(* IEC 61131-3 sources: volt/packages/volt-lsp-iec/test-corpus/bakon-nano/Device/Plc Logic/Application/Library Manager/L_EtcSlaveConfig, 51 files *)

(* ---- _L_ECC_ESCHEDULE.dut ---- *)
TYPE _L_ECC_ESCHEDULE :
(
	INIT := 0,
	INIT_DONE := 99,
	SCHEDULING_ACTIVE := 10
);
END_TYPE

(* ---- _L_ECC_ESEVERITY.dut ---- *)
TYPE _L_ECC_ESEVERITY :
(
	NO_RESPONSE := 0,
	WARNING := 2,
	INFORMATION := 11,
	WARNING_LOCK := 13,
	FAULT_LOG := 18,
	FAULT_QSPAPPL := 19,
	FAULT_QSP := 20,
	FAULT_QSP_CINH := 21,
	FAULT_CINH := 23,
	FAULT := 30
);
END_TYPE

(* ---- _L_ECC_ESTEPPER.dut ---- *)
TYPE _L_ECC_ESTEPPER :
(
	INIT := 0,
	INIT_DONE := 99,
	READ_IDENTITY_INIT := 10,
	READ_IDENTITY_DEVICENAME,
	READ_IDENTITY_HARDWAREVERSION,
	READ_IDENTITY_SOFTWAREVERSION,
	READ_IDENTITY_SYSTEMVERSION,
	READ_IDENTITY_VENDORID,
	READ_IDENTITY_PRODUCTCODE,
	READ_IDENTITY_REVISION,
	READ_IDENTITY_SERIALNUMBER,
	READ_IDENTITY_MANUFACTURER,
	READ_IDENTITY_DEVICECLASS,
	READ_IDENTITY_PRODUCTCODE_CD,
	READ_IDENTITY_FINISH_CD,
	C250_INIT := 100,
	C250_ERROR_REGISTER := 110,
	C250_CHECK_READING_REQUIRED,
	C250_EXTERNAL_TEMPERATURE := 115,
	C250_STATE_INPUTS,
	C250_STATE_OUTPUTS,
	C250_CPU1_REFERENCE_VOLTAGE := 120,
	C250_CPU1_24V_VOLTAGE := 121,
	C250_CPU1_5V_VOLTAGE := 122,
	C250_CPU1_3V3_VOLTAGE := 123,
	C250_CPU1_TEMPERATURE := 124,
	C250_CPU1_OUTPUT_CURRENT := 125,
	C250_CPU1_CYCLETIME := 126,
	C250_CPU1_ERROR_CODE := 127,
	C250_CPU1_ERROR_LINE := 128,
	C250_CPU1_ERROR_MODULE := 129,
	C250_CPU1_ERROR_CLASS := 130,
	C250_CPU1_ERROR_WRITETOCONTROLLER := 131,
	C250_CPU1_ERROR_WRITETOFRAMEWORK := 132,
	C250_CPU2_REFERENCE_VOLTAGE := 140,
	C250_CPU2_24V_VOLTAGE,
	C250_CPU2_5V_VOLTAGE,
	C250_CPU2_3V3_VOLTAGE,
	C250_CPU2_TEMPERATURE,
	C250_CPU2_OUTPUT_CURRENT,
	C250_CPU2_CYCLETIME,
	C250_CPU2_ERROR_CODE,
	C250_CPU2_ERROR_LINE,
	C250_CPU2_ERROR_MODULE,
	C250_CPU2_ERROR_CLASS,
	C250_CPU2_ERROR_WRITETOCONTROLLER,
	C250_CPU2_ERROR_WRITETOFRAMEWORK := 152,
	C250_DONE_WRITETOLOGS := 198,
	C250_DONE := 199,
	S13X_INIT := 200,
	S13X_DISABLE_AUTO_ACK,
	S13X_ERROR_REGISTER_HARDWARE := 210,
	S13X_ERROR_REGISTER_DIAGNOSTIC,
	S13X_MODULE_STATUS_DIAGNOSTIC,
	S13X_CHECK_READING_REQUIRED,
	S13X_COUPLER_VERSION_FPGA := 220,
	S13X_COUPLER_VERSION_BACKPLANE,
	S13X_COUPLER_VERSION_FIRMWARE,
	S13X_COUPLER_MX_FILE,
	S13X_COUPLER_NUMBER_OF_SLICES,
	S13X_SLICE_INIT := 230,
	S13X_SLICE_VERSION_FPGA,
	S13X_SLICE_VERSION_MODULE,
	S13X_SLICE_SERIALNUMBER,
	S13X_SLICE_MX_FILE,
	S13X_SLICE_ID_CONFIGURED,
	S13X_SLICE_ADDRESS,
	S13X_SLICE_ID_DETECTED,
	S13X_SLICE_DONE,
	S13X_SLICE_SW_VERSION,
	S13X_SLICE_HW_VERSION,
	S13X_SLICE_MODULE_ID,
	S13X_SLICE_ERROR_HARDWARE_SLOT := 250,
	S13X_SLICE_ERROR_HARDWARE_DIAG1,
	S13X_SLICE_ERROR_HARDWARE_DIAG2,
	S13X_SLICE_ERROR_HARDWARE_DIAG3,
	S13X_SLICE_ERROR_HARDWARE_DIAG4,
	S13X_SLICE_ERROR_HARDWARE_WRITE_ACK,
	S13X_SLICE_ERROR_HARDWARE_WRITETOCONTROLLER,
	S13X_SLICE_ERROR_HARDWARE_WRITETOFRAMEWORK,
	S13X_SLICE_ERROR_DIAGNOSTIC_READSLOT,
	S13X_SLICE_ERROR_DIAGNOSTIC_WRITESLOT,
	S13X_SLICE_ERROR_DIAGNOSTIC_DIAG1,
	S13X_SLICE_ERROR_DIAGNOSTIC_DIAG2,
	S13X_SLICE_ERROR_DIAGNOSTIC_DIAG3,
	S13X_SLICE_ERROR_DIAGNOSTIC_DIAG4,
	S13X_SLICE_ERROR_DIAGNOSTIC_WRITE_ACK,
	S13X_SLICE_ERROR_DIAGNOSTIC_WRITETOCONTROLLER,
	S13X_SLICE_ERROR_DIAGNOSTIC_WRITETOFRAMEWORK,
	S13X_DONE_WRITETOLOGS := 298,
	S13X_DONE := 299,
	ISERIES_INIT := 400,
	ISERIES_STEP_1 := 401,
	ISERIES_STEP_2 := 402,
	ISERIES_STEP_3 := 403,
	ISERIES_STEP_4 := 404,
	ISERIES_STEP_5 := 405,
	ISERIES_DONE := 499
);
END_TYPE

(* ---- FILE_STATE.dut ---- *)
TYPE FILE_STATE :
(
	S_NONE,
	S_INITIALIZE,
	S_GET_SLAVE_STATE,
	S_WAIT_FILE_SIZE,
	S_WAIT_FILE_OPEN,
	S_READ_FILE,
	S_CLOSE_FILE,
	S_PROCESS,
	S_READ_PAR_RECORDS,
	S_WAIT_XFER_COMPLETE,
	S_ERROR,
	S_DONE
);
END_TYPE

(* ---- L_ECC_EC250_CPUNUMBER.dut ---- *)
TYPE L_ECC_EC250_CPUNUMBER :
(
	NO_CPU := 0,
	CPU_1 := 1,
	CPU_2 := 2,
	CPU_3 := 3
);
END_TYPE

(* ---- L_ECC_EC250_ERRORCLASS.dut ---- *)
TYPE L_ECC_EC250_ERRORCLASS :
(
	NO_ERROR := 0,
	SYNCHRONIZATION_ERROR := 1,
	COMMUNICATION_ERROR := 2,
	IO_ERROR := 3,
	ERRORHANDLER_ERROR := 4,
	FATAL_ERROR := 5
);
END_TYPE

(* ---- L_ECC_EC250_ERRORCODE.dut ---- *)
TYPE L_ECC_EC250_ERRORCODE :
(
	OK := 0,
	HWT_PARAMETER_ERROR := 1,
	HWT_INIT_ERROR := 2,
	HWT_MEM_MARCHC_ERROR := 100,
	HWT_MEM_GALPAT_ERROR := 101,
	HWT_STACK_UNDERFLOW_ERROR := 200,
	HWT_STACK_OVERFLOW_ERROR := 201,
	HWT_CPU_ERROR := 300,
	WT_FW_ERROR := 400,
	HWT_FWINTERFACE_ERROR := 500,
	HWT_ADC_ERROR := 504,
	HWT_DMA_ERROR := 505,
	HWT_CRC_ERROR := 506,
	HWT_TIMER_ERROR := 507,
	HWT_CLOCK_ERROR := 508,
	HWT_SOFTERROR := 509,
	HWT_DIVZERO := 510,
	TIMEOUT_ERR := 512,
	OUT_OF_RANGE_ERR := 513,
	OVERWRITE_ERR := 514,
	UNDERFLOW_ERR := 515,
	PRG_CNTRL_ERR := 516,
	INIT_ERROR := 528,
	ASSERT_TRUE_ERR := 592,
	ASSERT_NOT_NULL_ERR := 593,
	ASSERT_GE_ERR := 594,
	ASSERT_GT_ERR := 595,
	ASSERT_LE_ERR := 596,
	ASSERT_LT_ERR := 597,
	ASSERT_NE_ERR := 598,
	ASSERT_EQ_ERR := 599,
	ASSERT_FALSE_ERR := 600,
	TP_OUT_NOT_SPECIFIED := 640,
	TP_OUT_NOT_RECOGNIZED := 641,
	TP_OUT_NOT_ACTIVE := 642,
	TP_INP_BUSY := 656,
	TP_INP_CROSSTALK := 657,
	TP_INP_NOT_RECOGNIZED := 658,
	TP_INTINP_NOT_RECOGNIZED := 659,
	TP_INP_LOST := 660,
	TP_INVALID_COUNT_FOR_SELECTOR := 661,
	MRAM_READ_ERR := 673,
	MRAM_WRITE_ERR := 674,
	MRAM_INDEX_OUT_OF_RANGE := 675,
	MRAM_CORRUPT_PAGE_SIZE := 676,
	MRAM_CRC_ERR := 677,
	MRAM_MAGICNUMBER_ERR := 678,
	RESET_LOW_POWER := 768,
	RESET_WINDOW_WD := 769,
	RESET_INDEPENDENT_WD := 770,
	RESET_SW := 771,
	RESET_POWER_ON_DOWN := 772,
	RESET_NMI := 773,
	RESET_BROWNOUT := 774,
	RESET_NO_REASON := 775,
	ADC_REF_LOW := 1024,
	ADC_REF_HIGH := 1025,
	ADC_24V_LOW := 1026,
	ADC_24V_HIGH := 1027,
	ADC_5V_LOW := 1028,
	ADC_5V_HIGH := 1029,
	ADC_3_3V_LOW := 1030,
	ADC_3_3V_HIGH := 1031,
	ADC_TEMP_LOW := 1032,
	ADC_TEMP_HIGH := 1033,
	ADC_CURR_HIGH := 1034,
	ADC_24V_FATAL := 1035,
	LINE_TIMEOUT := 1280,
	NOVALIDCPUID := 1281,
	TIMEOUTTIMERERR := 1282,
	DIPSWITCHREADERR := 1283,
	DIPSWITCHCHANGED := 1284,
	DIPSWITCHXCHGERROR := 1285,
	DIPSWITCH_INVALID_ADDRESS := 1286,
	CLK_ERROR := 1312,
	CLK_PARTNER_LOW := 1313,
	CLK_PARTNER_HIGH := 1314,
	HW_REVISION_ERROR := 1328,
	INPUTXCHGERROR := 1536,
	INPUT_TIMEOUT := 1537,
	INPUT_EXTMATTE_KS := 1552,
	INPUT_EXTMATTE_OPEN := 1553,
	OUTPUTXCHGERROR := 1792,
	OUTPUTFAIL := 1793,
	OUTPUT_WAITFB := 1794,
	OUTPUT_TIMEOUT := 1795,
	OUTPUT_HSTP_TIMEOUT := 1796,
	OUTPUT_LSTP_TIMEOUT := 1797,
	OUTPUT_LSTP_CONNECT_ERR := 1798,
	OUTPUT_USTP_TIMEOUT := 1799,
	OUTPUT_NOPAR_USED := 1800,
	BCOM_NOTREADY := 2048,
	BCOM_BUSY := 2049,
	BCOM_NONEWDATA := 2050,
	BCOM_CRCERR := 2051,
	BCOM_BITERR := 2052,
	XCOM_NOTREADY := 2304,
	XCOM_BUSY := 2305,
	XCOM_NONEWDATA := 2306,
	XCOM_CRCERR := 2307,
	I2C_TIMEOUT := 2560,
	I2C_BUSY := 2561,
	FSOE_RESET_IND := 2816,
	FSOE_INVALID_CMD := 2817,
	FSOE_UNKNOWN_CMD := 2818,
	FSOE_INVALID_CONNID := 2819,
	FSOE_INVALID_CRC := 2820,
	FSOE_WD_EXPIRED := 2821,
	FSOE_INVALID_ADDRESS := 2822,
	FSOE_INVALID_DATA := 2823,
	FSOE_INVALID_COMMPARALEN := 2824,
	FSOE_INVALID_COMMPARA := 2825,
	FSOE_INVALID_USERPARALEN := 2826,
	FSOE_INVALID_USERPARA := 2827,
	FSOE_INVALID_TP_INP_DURATION := 2828,
	FSOE_INVALID_TP_INP_FREQUENCY := 2829,
	FSOE_INVALID_TP_OUT_DURATION := 2830,
	FSOE_INVALID_TP_OUT_FREQUENCY := 2831,
	FSOE_INVALID_WATCHDOG_TIME := 2832,
	FSOE_INVALID_INP_EXT_SUPPLY := 2833,
	FSOE_INVALID_INP_IN_USE := 2834,
	FSOE_INVALID_INP_USED_EXT_MISMATCH := 2835,
	FSOE_INVALID_OUT_IN_USE := 2836,
	FSOE_INVALID_OUT_USED_EXT_MISMATCH := 2837,
	FSOE_EXTENDED_ERROR := 2944,
	FSOE_ERROR := 2992,
	TH_GLOBAL_ERROR := 3072,
	TH_TIMEOUT := 3073,
	MC1_ID_INVALID := 3329,
	MC2_ID_INVALID := 3330,
	MC3_ID_INVALID := 3331,
	FOREIGN_ERROR_DETECTED := 3584,
	FLASH_TIMEOUT := 3841,
	FLASH_LOCKED := 3842,
	FLASH_BUSY := 3851,
	FLASH_ERROR := 3854
);
END_TYPE

(* ---- L_ECC_EC250_ERRORMODULE.dut ---- *)
TYPE L_ECC_EC250_ERRORMODULE :
(
	OBJ_UNKNOWN_ID := 0,
	OBJ_FSOETASK_ID := 4,
	OBJ_INPUT_ID := 8,
	OBJ_MAINTASK_ID := 12,
	OBJ_PRGCONTRLTASK_ID := 16,
	OBJ_SYNCSAFETYPARTNER_ID := 20,
	OBJ_XCOM_ID := 24,
	OBJ_SAFETYHAL_ID := 28,
	OBJ_YSTIMER_ID := 32,
	OBJ_MSTIMER_ID := 36,
	OBJ_BASEBOARDCOM_ID := 44,
	OBJ_DIPSWITCH_ID := 48,
	OBJ_HELPER_ID := 52,
	OBJ_SYNCLINE_ID := 56,
	OBJ_TIMETABLE_ID := 60,
	OBJ_TESTHANDLER_ID := 64,
	OBJ_TIME_ITERATOR_ID := 80,
	OBJ_SPI_ID := 96,
	OBJ_TIMER_ID := 97,
	OBJ_BACKUPSRAM_ID := 98,
	OBJ_PWR_ID := 99,
	OBJ_RCC_ID := 100,
	OBJ_GPIO_ID := 101,
	OBJ_DMASTREAM_ID := 102,
	OBJ_ADC_ID := 103,
	OBJ_WD_ID := 104,
	OBJ_FLASH_ID := 105,
	OBJ_I2C_ID := 106,
	OBJ_INPUTHANDLER_ID_1 := 128,
	OBJ_INPUTHANDLER_ID_2 := 129,
	OBJ_INPUTHANDLER_ID_3 := 130,
	OBJ_INPUTHANDLER_ID_4 := 131,
	OBJ_OUTPUT_ID_1 := 144,
	OBJ_OUTPUT_ID_2 := 145,
	OBJ_USTESTPULSE_ID := 148,
	OBJ_OUTPUTHANDLER_ID := 160,
	OBJ_OUTPFSWITCH_ID := 164
);
END_TYPE

(* ---- L_ECC_EDEVICETYPE.dut ---- *)
TYPE L_ECC_EDEVICETYPE :
(
	UNKNOWN := 0,
	C25BAYCB := 16#43004342,
	C25BAYSQ := 16#43005153,
	C25BAYA42 := 16#43000402,
	C25BAYA82 := 16#43000802,
	C25BAYA160 := 16#43001000,
	C25BAYA164 := 16#43001004,
	EPM_S130 := 16#514,
	EPM_S131 := 16#51E,
	EPM_S200 := 16#19F82,
	EPM_S201 := 16#39F84,
	EPM_S202 := 16#59FC1,
	EPM_S203 := 16#89F84,
	EPM_S204 := 16#29F82,
	EPM_S205 := 16#49F84,
	EPM_S206 := 16#79FC1,
	EPM_S207 := 16#F0147C1,
	EPM_S208 := 16#F0347C2,
	EPM_S209 := 16#139FC1,
	EPM_S210 := 16#121F41,
	EPM_S300 := 16#101AF90,
	EPM_S301 := 16#104AFA0,
	EPM_S302 := 16#106AFC8,
	EPM_S303 := 16#103AF90,
	EPM_S304 := 16#105AFA0,
	EPM_S305 := 16#107AFC8,
	EPM_S306 := 16#102AF90,
	EPM_S308 := 16#109AF90,
	EPM_S309 := 16#108AFA0,
	EPM_S310 := 16#F4157E1,
	EPM_S311 := 16#F4357E2,
	EPM_S312 := 16#1132F48,
	EPM_S400 := 16#40115C3,
	EPM_S401 := 16#40415C4,
	EPM_S402 := 16#40215C3,
	EPM_S403 := 16#40515C4,
	EPM_S404 := 16#4061544,
	EPM_S405 := 16#4031543,
	EPM_S406 := 16#40C1543,
	EPM_S408 := 16#40B1543,
	EPM_S409 := 16#4111543,
	EPM_S410 := 16#40715C3,
	EPM_S411 := 16#8411809,
	EPM_S412 := 16#40D1544,
	EPM_S413 := 16#4121544,
	EPM_S414 := 16#40E1544,
	EPM_S415 := 16#40F1543,
	EPM_S416 := 16#8842880,
	EPM_S500 := 16#50125D8,
	EPM_S501 := 16#50325E0,
	EPM_S502 := 16#50225D8,
	EPM_S503 := 16#50425E0,
	EPM_S504 := 16#50B25D8,
	EPM_S505 := 16#50A25E0,
	EPM_S600 := 16#8C13800,
	EPM_S601 := 16#8C3380A,
	EPM_S602 := 16#8C23801,
	EPM_S603 := 16#8C4388B,
	EPM_S604 := 16#9C17800,
	EPM_S606 := 16#8812880,
	EPM_S620 := 16#9014880,
	EPM_S640 := 16#E010700,
	EPM_S650 := 16#E411700
);
END_TYPE

(* ---- L_ECC_EEPMSXXX_ERRORCODE.dut ---- *)
TYPE L_ECC_EEPMSXXX_ERRORCODE :
(
	OK := 0,
	INTERNAL_ERROR := 1,
	EXTERNAL_ERROR := 2,
	CHANNEL_ERROR := 3,
	SUPPLY_VOLTAGE_ERROR := 4,
	PARAMETER_ERROR := 5,
	INTERNAL_COM_FAULT := 6,
	PROCESS_ALARM_LOST := 7,
	BROKEN_WIRE := 8,
	MEASURING_RANGE_UNDERFLOW := 9,
	MEASURING_RANGE_OVERFLOW := 10,
	LOST_OVERFLOW_UNDERFLOW_ALARM := 11,
	LOST_COMPARE_VALUE_RACHED_ALARM := 12,
	AUTO_ACK_DISABLED := 100
);
END_TYPE

(* ---- L_ECC_EERROR.dut ---- *)
TYPE L_ECC_EERROR :
(
	NOERROR := 0,
	NOSLAVECONNECTED,
	INVALIDSLAVECONNECTED,
	SLAVENOTREADYFORSDO,
	INVALIDSTATEMACHINE,
	INVALIDSLICENUMBER,
	COULDNOTSENDAUTOACKERROR,
	COULDNOTSENDDIAGNOSTICERROR
);
END_TYPE

(* ---- L_ECC_EEXTENDEDSTATE.dut ---- *)
TYPE L_ECC_EEXTENDEDSTATE :
(
	NONE := 16#0,
	INITIALIZING := 16#1,
	PREOPERATIONAL := 16#2,
	BOOTSTRAP := 16#3,
	SAFEOPERATIONAL := 16#4,
	OPERATIONAL := 16#8,
	UNKNOWN := 16#FFEF,
	FIRMWAREDOWNLOAD := 16#201,
	CABLENOTCONNECTED := 16#202,
	BUSMISMATCH := 16#203,
	CONNECTIONFAULTY := 16#801,
	NOTALLSLAVESOPERATIONAL := 16#802,
	CONNECTIONLOST := 16#803
);
END_TYPE

(* ---- L_ECC_SCC250_CPU.dut ---- *)
TYPE L_ECC_SCC250_CPU :
STRUCT
	ECPUNUMBER : L_ECC_eC250_CpuNumber;
	XERRORACTIVE : BOOL;
	EERRORCLASS : L_ECC_eC250_ErrorClass;
	EERRORCODE : L_ECC_eC250_ErrorCode;
	EPREVIOUSERRORCODE : L_ECC_eC250_ErrorCode;
	EERRORMODULE : L_ECC_eC250_ErrorModule;
	WERRORLINE : WORD;
END_STRUCT
END_TYPE

(* ---- L_ECC_SCDEVICEINFO.dut ---- *)
TYPE L_ECC_SCDEVICEINFO :
STRUCT
	UIDEVICEADDRESS : UINT;
	EDEVICETYPE : L_ECC_eDeviceType := L_ECC_eDeviceType.Unknown;
	SDEVICENAME : STRING(255);
	SHARDWAREVERSION : STRING(64);
	SSOFTWAREVERSION : STRING(64);
	USISYSTEMVERSION : USINT;
	DWVENDORID : DWORD;
	DWPRODUCTCODE : DWORD;
	DWREVISION : DWORD;
	DWSERIALNUMBER : DWORD;
END_STRUCT
END_TYPE

(* ---- L_ECC_SCEMPSXXX_DIAGNOSTIC.dut ---- *)
TYPE L_ECC_SCEMPSXXX_DIAGNOSTIC :
UNION
	SCEPMS404_S405 : L_ECC_scEPMS404_S405_Diagnostic;
	SCEPMS600 : L_ECC_scEPMS600_Diagnostic;
	SCEPMS601_S602 : L_ECC_scEPMS603_S604_Diagnostic;
	SCEPMS603_S604 : L_ECC_scEPMS603_S604_Diagnostic;
	SCGENERIC : L_ECC_scEMPSxxx_DiagnosticBits;
	ABYBYTES : ARRAY [1..4] OF BYTE;
	DWVALUE : DWORD;
END_UNION
END_TYPE

(* ---- L_ECC_SCEMPSXXX_DIAGNOSTICBITS.dut ---- *)
TYPE L_ECC_SCEMPSXXX_DIAGNOSTICBITS :
STRUCT
	BERROR : BIT;
	BINTERNALERROR : BIT;
	BEXTERNALERROR : BIT;
	BCHANNELERROR : BIT;
	BSUPPLYVOLTAGEERROR : BIT;
	BRESERVED_0 : BIT;
	BRESERVED_1 : BIT;
	BPARAMETERERROR : BIT;
	BRESERVED_2 : BIT;
	BRESERVED_3 : BIT;
	BRESERVED_4 : BIT;
	BRESERVED_5 : BIT;
	BINTERNALCOMFAULT : BIT;
	BRESERVED_6 : BIT;
	BPROCESSALARMLOST : BIT;
	BRESERVED_7 : BIT;
END_STRUCT
END_TYPE

(* ---- L_ECC_SCEPMS404_S405_DIAGNOSTIC.dut ---- *)
TYPE L_ECC_SCEPMS404_S405_DIAGNOSTIC :
STRUCT
	SCGENERAL : L_ECC_scEMPSxxx_DiagnosticBits;
	SCCHANNEL_0 : L_ECC_scEPMS404_S405_DiagnosticBits;
	SCCHANNEL_1 : L_ECC_scEPMS404_S405_DiagnosticBits;
END_STRUCT
END_TYPE

(* ---- L_ECC_SCEPMS404_S405_DIAGNOSTICBITS.dut ---- *)
TYPE L_ECC_SCEPMS404_S405_DIAGNOSTICBITS :
STRUCT
	BPARAMETERERROR : BIT;
	BRESERVED_0 : BIT;
	BRESERVED_1 : BIT;
	BRESERVED_2 : BIT;
	BBROKENWIRE : BIT;
	BPROCESSALARMLOST : BIT;
	BMEASURINGRANGEUNDERFLOW : BIT;
	BMEASURINGRANGEOVERFLOW : BIT;
END_STRUCT
END_TYPE

(* ---- L_ECC_SCEPMS600_DIAGNOSTIC.dut ---- *)
TYPE L_ECC_SCEPMS600_DIAGNOSTIC :
STRUCT
	SCGENERAL : L_ECC_scEMPSxxx_DiagnosticBits;
	SCCHANNEL_0 : L_ECC_scEPMS600_DiagnosticBits;
	BYRESERVED_1 : BYTE;
END_STRUCT
END_TYPE

(* ---- L_ECC_SCEPMS600_DIAGNOSTICBITS.dut ---- *)
TYPE L_ECC_SCEPMS600_DIAGNOSTICBITS :
STRUCT
	BHW_GATEOPENED : BIT;
	BHW_GATECLOSED : BIT;
	BENDVALUEOVERFLOWUNDERFLOW : BIT;
	BCOMPAREVALUEREACHED : BIT;
	BLATCHED : BIT;
	BRESERVED_0 : BIT;
	BRESERVED_1 : BIT;
	BRESERVED_2 : BIT;
END_STRUCT
END_TYPE

(* ---- L_ECC_SCEPMS601_S602_DIAGNOSTICBITS.dut ---- *)
TYPE L_ECC_SCEPMS601_S602_DIAGNOSTICBITS :
STRUCT
	BRESERVED_0 : BIT;
	BLOSTOVERFLOWUNDERFLOWALARM : BIT;
	BLOSTCOMPAREVALUEREACHEDALARM : BIT;
	BRESERVED_1 : BIT;
	BRESERVED_2 : BIT;
	BRESERVED_3 : BIT;
	BRESERVED_4 : BIT;
END_STRUCT
END_TYPE

(* ---- L_ECC_SCEPMS603_S604_DIAGNOSTIC.dut ---- *)
TYPE L_ECC_SCEPMS603_S604_DIAGNOSTIC :
STRUCT
	SCGENERAL : L_ECC_scEMPSxxx_DiagnosticBits;
	BYRESERVED_0 : BYTE;
	BYRESERVED_1 : BYTE;
END_STRUCT
END_TYPE

(* ---- L_ECC_SCS13X_COUPLER.dut ---- *)
TYPE L_ECC_SCS13X_COUPLER :
STRUCT
	WNUMBEROFIOSLICES : WORD;
	UIVERSION_FPGA : UINT;
	UIVERSION_BACKPLANE : UINT;
	UDIVERSION_FIRMWARE : UDINT;
	SMX_FILE : STRING(16);
END_STRUCT
END_TYPE

(* ---- L_ECC_SCS13X_IO_SLICE.dut ---- *)
TYPE L_ECC_SCS13X_IO_SLICE :
STRUCT
	EDEVICETYPE : L_ECC_eDeviceType := L_ECC_eDeviceType.Unknown;
	UDIVERSION_FPGA : UDINT;
	UDIVERSION_MODULE : UDINT;
	SSERIALNUMBER : STRING(22);
	SMX_FILE : STRING(16);
	UDICONFIGUREDID : UDINT;
	UDIDETECTEDID : UDINT;
	UIDETECTEDADDRESS : UINT;
	ABYDIAGNOSTICDATA : ARRAY [0..7] OF BYTE;
	PSCIOSLICE : POINTER TO L_IOSlice;
END_STRUCT
END_TYPE

(* ---- L_ECC_SCSCHEDULEDATA.dut ---- *)
TYPE L_ECC_SCSCHEDULEDATA :
STRUCT
	PFBINSTANCE : POINTER TO _L_ECC_XXX_Diagnostics;
END_STRUCT
END_TYPE

(* ---- L_ECC_SCSLAVESTATUS.dut ---- *)
TYPE L_ECC_SCSLAVESTATUS :
STRUCT
	SNAME : STRING;
	UIADDRESS : UINT;
	XPRESENT : BOOL;
	XOPTIONAL : BOOL;
	XOPERATIONAL : BOOL;
	EOPERATINGMODE : L_ECC_eExtendedState := L_ECC_eExtendedState.None;
	SCEMERGENCYMESSAGE : L_ETC_COE_EMERGENCY;
	UDIERRORCOUNT_IN : UINT;
	UDIERRORCOUNT_OUT : UINT;
END_STRUCT
END_TYPE

(* ---- PARAUPLOAD_STATE.dut ---- *)
TYPE PARAUPLOAD_STATE :
(
	UPL_INITIALIZE,
	UPL_WAIT_GET_SLAVE_STATE,
	UPL_UPLOADING,
	UPL_ERROR,
	UPL_DONE
);
END_TYPE

(* ---- L_ECC_INTERNAL.gvl ---- *)
VAR_GLOBAL
	SMANUFACTURER : STRING := 'Lenze';
	SDEVCLASSINV : STRING := 'Inverter';
END_VAR

(* ---- GETBOOLEANPROPERTY.pou ---- *)
FUNCTION GETBOOLEANPROPERTY : BOOL
VAR_INPUT
	STKEY : WSTRING;
END_VAR
END_FUNCTION

(* ---- GETCOMPANY.pou ---- *)
FUNCTION GETCOMPANY : WSTRING
END_FUNCTION

(* ---- GETNUMBERPROPERTY.pou ---- *)
FUNCTION GETNUMBERPROPERTY : DINT
VAR_INPUT
	STKEY : WSTRING;
END_VAR
END_FUNCTION

(* ---- GETTEXTPROPERTY.pou ---- *)
FUNCTION GETTEXTPROPERTY : WSTRING
VAR_INPUT
	STKEY : WSTRING;
END_VAR
END_FUNCTION

(* ---- GETTEXTPROPERTY2.pou ---- *)
FUNCTION GETTEXTPROPERTY2 : POINTER TO WSTRING
VAR_INPUT
	STKEY : WSTRING;
END_VAR
END_FUNCTION

(* ---- GETTITLE.pou ---- *)
FUNCTION GETTITLE : WSTRING
END_FUNCTION

(* ---- GETVERSION.pou ---- *)
FUNCTION GETVERSION : VERSION
END_FUNCTION

(* ---- GETVERSIONPROPERTY.pou ---- *)
FUNCTION GETVERSIONPROPERTY : VERSION
VAR_INPUT
	STKEY : WSTRING;
END_VAR
END_FUNCTION

(* ---- L_ECC_INITCDFORLENZEINVERTER.pou ---- *)
FUNCTION L_ECC_INITCDFORLENZEINVERTER : BOOL
VAR_INPUT
	PETCSLAVE : POINTER TO ETCSlave;
END_VAR
END_FUNCTION

(* ---- _L_ECC_XXX_DIAGNOSTICS.pou ---- *)
FUNCTION_BLOCK _L_ECC_XXX_DIAGNOSTICS
VAR_INPUT
	XENABLE : BOOL := TRUE;
END_VAR
VAR_OUTPUT
	XBUSY : BOOL;
	XDONE : BOOL;
	XDIAGACTIVE : BOOL;
	XERRORDETECTED : BOOL;
	XERROR : BOOL;
	EERRORID : L_ECC_eError;
END_VAR
VAR
	XBUSY_INT : BOOL := FALSE;
	XDONE_INT : BOOL := FALSE;
	XERROR_INT : BOOL := FALSE;
	EERRORID_INT : L_ECC_eError;
	XDIAGACTIVE_INT : BOOL := FALSE;
	XERRORDETECTED_INT : BOOL := FALSE;
	SCDEVICEINFO_INT : L_ECC_scDeviceInfo;
	PETCSLAVE_INT : POINTER TO L_ETC.ETCSlave;
	PETCSLAVE_MEM : POINTER TO L_ETC.ETCSlave;
	ESTEPPER : _L_ECC_eStepper;
	UIFORLOOP : UINT;
	XINITDONE : BOOL := FALSE;
	ECMASTER : POINTER TO L_IODrvEtherCAT;
	WMASTERSTATE : L_ETC_STATE := L_ETC_STATE.ETC_STATE_NONE;
	FBGETSLAVESTATE : L_ETC_GetSlaveState;
	WSLAVESTATE : L_ETC_STATE := L_ETC_STATE.ETC_STATE_NONE;
	XSDOSTOPONERROR : BOOL := TRUE;
	FBSDOREAD : L_ETC_CoE_SdoRead;
	FBSDOREAD_XEXECUTE_MEM : BOOL;
	ABYSDOREADRAWVALUES : ARRAY [0..uiSdoReadArraySize] OF BYTE;
	SSDOREADPARSEDVALUE : STRING(255);
	DWSDOREADPARSEDVALUE : DWORD;
	FBSDOWRITE : L_ETC_CoE_SdoWrite;
	ABYSDOWRITERAWVALUES : ARRAY [0..uiSdoWriteArraySize] OF BYTE;
	XSDO_READSYSTEMVERSION : BOOL;
	XFIRSTCALL : BOOL := TRUE;
	XREADCOMPONENTINFODONE : BOOL;
	UISDOREADARRAYSIZE : UINT := 127;
	UISDOWRITEARRAYSIZE : UINT := 3;
	UDISDOTIMEOUT : UDINT := 1000;
END_VAR
END_FUNCTION_BLOCK

METHOD GETDEVICECLASS : BOOL
VAR_IN_OUT
	SDEVICECLASS : STRING;
END_VAR
END_METHOD

METHOD INITFIRSTCALL
END_METHOD

METHOD SETCMPINFODATA : BOOL
END_METHOD

METHOD AMAIN
END_METHOD

METHOD ASTATEMACHINE
END_METHOD

METHOD MCHECKDEVICETYPE : BOOL
VAR_INPUT
	DWPRODUCTID : DWORD;
END_VAR
END_METHOD

METHOD MRESETOUTPUTS
END_METHOD

METHOD MSDO_READ : BOOL
VAR_INPUT
	WINDEX : WORD;
	BYSUBINDEX : BYTE;
END_VAR
END_METHOD

METHOD MSDO_WRITE : BOOL
VAR_INPUT
	WINDEX : WORD;
	BYSUBINDEX : BYTE;
	BYSIZE : BYTE;
	DWVALUE : DWORD;
END_VAR
END_METHOD

METHOD MSETETCSLAVE : BOOL
VAR_INPUT
	PETCSLAVE : POINTER TO ETCSlave;
END_VAR
END_METHOD

(* ---- ETCCONFIGPARAXFER.pou ---- *)
FUNCTION_BLOCK ETCCONFIGPARAXFER EXTENDS L_SUDP_UpDownload
VAR_INPUT
	XPREVENTETCOPERATIONALWHENSDOWRITEERROR : BOOL;
END_VAR
VAR
	BYOLDVALUEOFCONTROLINPUT : BYTE := 16#FF;
	WPARAFILESZ : INT;
	INUMBYTESIO : INT;
	IBUFOFFSET : INT;
	BHEADERTEST : BOOL;
	BIOABORTED : BOOL;
	STATE : FILE_STATE := S_INITIALIZE;
	SPARAFILENAME : STRING(255);
	HPARAFILE : CAA.HANDLE;
	ELASTERROR : L_SUDP_ErrorCodes;
	IPARDATASZ : INT;
	IPARRECSZ : INT;
	FGETFS : FILE.GetSize;
	FOPEN : FILE.Open;
	FREAD : FILE.Read;
	FCLOSE : FILE.Close;
	PIOBUFFER : POINTER TO BYTE;
	AYIOBUFFER : ARRAY [0..1000] OF BYTE;
	PPARMREC : POINTER TO L_SUDP_PARM_RECORD;
	PFILEHDR : POINTER TO L_SUDP_PAR_FILE_HDR;
	PPARMDAT : POINTER TO L_SUDP_PAR_DATA_HDR;
	PETCDEV : POINTER TO ETCSlave;
	ECONTROL : L_SUDP_Control;
	PSATTACHEDERRORTXT : POINTER TO STRING;
	SDOWR : L_ETC_CoE_SdoWrite;
	BIGNOREPARAMETER : BOOL;
	BSDOWRITEERROROCCURS : BOOL;
	GETSLAVESTATE : L_ETC_GetSlaveState;
	GETETCMASTERDIAGNOSTIC : L_ETC_GetMasterDiagnostic;
END_VAR
END_FUNCTION_BLOCK

METHOD CLOSEFILE
END_METHOD

METHOD DOWNLOAD
END_METHOD

METHOD IGNOREINDEX : BOOL
VAR_INPUT
	U16INDEX : UINT;
	U16SUBINDEX : UINT;
END_VAR
END_METHOD

METHOD INITIALIZE
VAR_INPUT
	PETCREMDEV : POINTER TO L_ETCSlave;
END_VAR
END_METHOD

METHOD RESETALLSIGNALS
END_METHOD

(* ---- ETCPARAMETERUPLOAD.pou ---- *)
FUNCTION_BLOCK ETCPARAMETERUPLOAD EXTENDS L_SUDP_UpDownload
VAR_INPUT
	DWFILEOFFSETCHECKSUMCALC : DWORD;
END_VAR
VAR
	PETCDEV : POINTER TO ETCSlave;
	ECONTROL : L_SUDP_Control;
	BYOLDVALUEOFCONTROLINPUT : BYTE := 16#FF;
	UPLSTATE : PARAUPLOAD_STATE := PARAUPLOAD_STATE.UPL_INITIALIZE;
	GETSLAVESTATE : L_ETC_GetSlaveState;
	GETETCMASTERDIAGNOSTIC : L_ETC_GetMasterDiagnostic;
	EUPLOADERROR : L_SUDP_ErrorCodes;
	PRMREADWRITEETC : L_SUDP_PRMFile_ReadWrite_ETC;
END_VAR
END_FUNCTION_BLOCK

METHOD INITIALIZE
VAR_INPUT
	PETCREMDEV : POINTER TO L_ETCSlave;
END_VAR
END_METHOD

METHOD PARAUPLOAD
END_METHOD

(* ---- GLOBALTEXTLIST.pou ---- *)
FUNCTION_BLOCK GLOBALTEXTLIST
VAR
	M_TEXTLISTFILE : STRING(255);
	_STNAMESPACE : STRING;
END_VAR
END_FUNCTION_BLOCK

(* ---- L_ECC_CD_DIAGNOSTIC.pou ---- *)
FUNCTION_BLOCK L_ECC_CD_DIAGNOSTIC EXTENDS _L_ECC_XXX_Diagnostics
VAR
	UIACTSLAVECOUNT : UINT := 0;
	UIACTSLAVEINPROGRESS : UINT;
	PSLAVES : ARRAY [1..uicMaxSlaves] OF POINTER TO ETCSlave;
	USISLAVESSTATE : ARRAY [1..uicMaxSlaves] OF USINT;
	XDATAUPDATED : BOOL;
	UICMAXDEPTH : UINT := 10;
	UICMAXSLAVES : UINT := 256;
END_VAR
END_FUNCTION_BLOCK

METHOD ADDSLAVE : BOOL
VAR_INPUT
	PECATSLAVE : POINTER TO ETCSlave;
END_VAR
END_METHOD

METHOD CHECKECATSLAVE : BOOL
VAR_INPUT
	PCHILD : POINTER TO IoConfigConnector;
END_VAR
END_METHOD

METHOD GETDATA : BOOL
VAR_INPUT
	COMPONENTINFOID : UDINT;
	NEXTSTEP : _L_ECC_eStepper;
END_VAR
VAR_IN_OUT
	STEPPER : _L_ECC_eStepper;
END_VAR
END_METHOD

METHOD UPDATECOMPONENTINFO : BOOL
VAR_INPUT
	DATASELECTION : UDINT;
	SDATA : STRING;
END_VAR
END_METHOD

METHOD AMAIN
END_METHOD

METHOD ASTATEMACHINE
END_METHOD

METHOD MCHECKDEVICETYPE : BOOL
VAR_INPUT
	DWPRODUCTID : DWORD;
END_VAR
END_METHOD

(* ---- L_ECC_S131_DIAGNOSTICS.pou ---- *)
FUNCTION_BLOCK L_ECC_S131_DIAGNOSTICS EXTENDS _L_ECC_XXX_Diagnostics
VAR
	SCBUSCOUPLER_INT : L_ECC_scS13x_Coupler;
	ASCIOSLICES_INT : ARRAY [1..uicMaxIOSlices] OF L_ECC_scS13x_IO_Slice;
	XSLICEREGISTERDONCMPDIR : BOOL;
	XSDO_READSLICESERIALNUMBER : BOOL;
	XSDO_READSLICEMXFILE : BOOL;
	WTEXTREFID : WORD;
	WSELECTEDIOSLICE : WORD;
	WRESETIOSLICES : WORD;
	DWERRORREGISTERHARDWARE_INT : DWORD;
	DWERRORREGISTERDIAGNOSTIC_INT : DWORD;
	LWMODULESTATUSDIAGNOSTIC_INT : DWORD;
	DWDISABLEAUTOACK_INT : DWORD;
	DWERRORCODEHARDWARE_INT : DWORD;
	DWERRORCODEDIAGNOSTIC_INT : DWORD;
	BYSLICEERRORSLICE_HARDWARE : BYTE;
	BYSLICEERRORSLICE_DIAGNOSTIC : BYTE;
	XHARDWAREERRORDETECTED_INT : BOOL := FALSE;
	XDIAGNOSTICERRORDETECTED_INT : BOOL := FALSE;
	SPRODUCTVERSION : STRING;
	SSERIALNUMBER : STRING;
	SHWVERSION : STRING;
	SSWVERSION : STRING;
	SMODULEID : STRING;
	UICMAXIOSLICES : UINT := 64;
END_VAR
END_FUNCTION_BLOCK

METHOD GETDEVICECLASS : BOOL
VAR_IN_OUT
	SDEVICECLASS : STRING;
END_VAR
END_METHOD

METHOD INITFIRSTCALL
END_METHOD

METHOD SETSLICECMPINFODATA : BOOL
END_METHOD

METHOD ACYCLICSTATEMACHINE
END_METHOD

METHOD AINITIALIZATIONSTATEMACHINE
END_METHOD

METHOD ASTATEMACHINE
END_METHOD

METHOD MCHECKDEVICETYPE : BOOL
VAR_INPUT
	DWPRODUCTID : DWORD;
END_VAR
END_METHOD

METHOD MCLEARIOSLICEREGISTRATIONS : BOOL
END_METHOD

METHOD MREGISTERIOSLICE : BOOL
VAR_INPUT
	PSCIOSLICE : POINTER TO L_IOSlice;
	BYSLOTNUMBER : BYTE;
END_VAR
END_METHOD

METHOD MRESETOUTPUTS
END_METHOD

METHOD MSETAUTOACKERROR : BOOL
END_METHOD

METHOD MSETDIAGNOSTICERROR : BOOL
VAR_INPUT
	BYSLICE : BYTE := 1;
	ESEVERITY : _L_ECC_eSeverity := _L_ECC_eSeverity.Fault_Log;
	DWERRORID : DWORD := 0;
END_VAR
END_METHOD

(* ---- L_ECC_SAFETY_DIAGNOSTICS.pou ---- *)
FUNCTION_BLOCK L_ECC_SAFETY_DIAGNOSTICS EXTENDS _L_ECC_XXX_Diagnostics
VAR
	SCCPU_1_INT : L_ECC_scC250_CPU;
	SCCPU_2_INT : L_ECC_scC250_CPU;
	XSDO_SLAVEISIOMODULE : BOOL;
	WTEXTREFID : WORD;
	DWERRORREGISTER_INT : DWORD;
	DWSTATEINPUT_MEM : DWORD;
	DWSTATEOUTPUT_MEM : DWORD;
	DWSTATEINPUT_INT : DWORD;
	DWSTATEOUTPUT_INT : DWORD;
	DWERRORCOUNT : DWORD;
	DWCLEARCOUNT : DWORD;
END_VAR
END_FUNCTION_BLOCK

METHOD GETDEVICECLASS : BOOL
VAR_IN_OUT
	SDEVICECLASS : STRING;
END_VAR
END_METHOD

METHOD ASTATEMACHINE
END_METHOD

METHOD MCHECKDEVICETYPE : BOOL
VAR_INPUT
	DWPRODUCTID : DWORD;
END_VAR
END_METHOD

METHOD MDECODESERIALNUMBER : STRING(11)
VAR_INPUT
	DWSERIALNUMBERBITCODED : DWORD;
END_VAR
END_METHOD

METHOD MRESETOUTPUTS
END_METHOD

METHOD MRESETOUTPUTS_ERRORS
END_METHOD

METHOD MSETDIAGNOSTICERROR : BOOL
VAR_INPUT
	ESEVERITY : _L_ECC_eSeverity := _L_ECC_eSeverity.Fault_Log;
	PSCCPUINFO : POINTER TO L_ECC_scC250_CPU;
END_VAR
END_METHOD

(* ---- L_ECC_SCHEDULER.pou ---- *)
FUNCTION_BLOCK L_ECC_SCHEDULER
VAR_INPUT
	XENABLE : BOOL := TRUE;
END_VAR
VAR
	HEVENTUPDATECONFIGURATIONDONE : RTS_IEC_HANDLE;
	HINTERFACEUPDATECONFIGURATIONDONE : RTS_IEC_HANDLE;
	ITFCALLBACK : CmpEventMgr.ICmpEventCallback;
	MYCONNECTOR : POINTER TO IoConfigConnector;
	SCHEDULER : L_ECC_XXX_Diagnostics_Scheduler;
	COMPONENTDIRECTORY : L_ECC_CD_Diagnostic;
	UICMAXDEPTH : UINT := 10;
END_VAR
END_FUNCTION_BLOCK

METHOD CHILDHASDIAGFB : BOOL
VAR_INPUT
	PCHILD : POINTER TO IoConfigConnector;
END_VAR
END_METHOD

METHOD CYCLICCALL : UDINT
END_METHOD

METHOD EVENTCALLBACK : UDINT
VAR_INPUT
	PEVENTPARAM : POINTER TO EventParam;
END_VAR
END_METHOD

METHOD FB_EXIT : BOOL
VAR_INPUT
	BINCOPYCODE : BOOL;
END_VAR
END_METHOD

METHOD FB_INIT : BOOL
VAR_INPUT
	BINITRETAINS : BOOL;
	BINCOPYCODE : BOOL;
END_VAR
END_METHOD

METHOD GETDIAGFBINSTANCE : POINTER TO _L_ECC_XXX_Diagnostics
VAR_INPUT
	PCHILD_ECATSLAVE : POINTER TO IoConfigConnector;
END_VAR
END_METHOD

METHOD GETDIAGSLAVES : BOOL
END_METHOD

METHOD GETDIAGSLAVESRECURSIVE : BOOL
VAR_INPUT
	PFATHER : POINTER TO IoConfigConnector;
	PCONNLIST : POINTER TO IoConfigConnector;
	CONNLISTCOUNT : DINT;
	DWDEPTH : DWORD;
END_VAR
END_METHOD

METHOD GETECATMASTECONNECTOR : BOOL
VAR_IN_OUT
	PECATMASTERCONNECTOR : POINTER TO IoConfigConnector;
END_VAR
END_METHOD

METHOD INITIALIZE : UDINT
VAR_INPUT
	WMODULETYPE : UINT;
	DWINSTANCE : UDINT;
	PCONNECTOR : POINTER TO IoConfigConnector;
END_VAR
END_METHOD

METHOD NODEISECATMASTER : BOOL
VAR_INPUT
	PNODE : POINTER TO IoConfigConnector;
END_VAR
END_METHOD

(* ---- L_ECC_XXX_DIAGNOSTICS_SCHEDULER.pou ---- *)
FUNCTION_BLOCK L_ECC_XXX_DIAGNOSTICS_SCHEDULER
VAR
	ASCHEDULEDATA : ARRAY [1..uicMaxFBs] OF L_ECC_scScheduleData;
	WNUMREGISTEREDFBS : WORD := 0;
	WMAXFBSPERCYCLE_INT : WORD := 1;
	UISCHEDULEIDX : UINT := 1;
	UISCHEDULELOOPCOUNT : UINT := 0;
	UISCHEDULELOOPMAX : UINT := 0;
	ESCHEDULER : _L_ECC_eSchedule := _L_ECC_eSchedule.INIT;
	DWDIAGCYCLECOUNT : DWORD := 0;
	DWDOUBLEREGISTRATIONCOUNT : DWORD := 0;
	UICMAXFBS : UINT := 256;
END_VAR
END_FUNCTION_BLOCK

METHOD AMAIN
END_METHOD

METHOD ASCHEDULE
END_METHOD

METHOD MFBISREGISTERED : BOOL
VAR_INPUT
	PFB_INSTANCE : POINTER TO _L_ECC_XXX_Diagnostics;
END_VAR
END_METHOD

METHOD MINIT : INT
VAR_INPUT
	WMAXFBSPERCYCLE : WORD := 1;
END_VAR
END_METHOD

METHOD MREGISTERFB : BOOL
VAR_INPUT
	PFB_INSTANCE : POINTER TO _L_ECC_XXX_Diagnostics;
END_VAR
END_METHOD

METHOD MSTOPSCHEDULING : BOOL
END_METHOD

(* ---- L_ETCSLAVE.pou ---- *)
FUNCTION_BLOCK L_ETCSLAVE
VAR_OUTPUT
	PETCSLAVE : POINTER TO ETCSlave;
END_VAR
VAR
	ETCSLAVE : ETCSlave;
	M_HLEMACCESS : RTS_IEC_HANDLE;
	PARSETXFER : EtcConfigParaXfer;
	PARSETUPLOAD : EtcParameterUpload;
	ISMANDATORY : BOOL;
	ISPRESENT : BOOL;
	MODULEHANDLER : L_IMHP_IModuleHandler;
END_VAR
END_FUNCTION_BLOCK

METHOD CYCLICCALL : UDINT
END_METHOD

METHOD FB_EXIT : BOOL
VAR_INPUT
	BINCOPYCODE : BOOL;
END_VAR
END_METHOD

METHOD FB_INIT : BOOL
VAR_INPUT
	BINITRETAINS : BOOL;
	BINCOPYCODE : BOOL;
END_VAR
END_METHOD

METHOD INITIALIZE : UDINT
VAR_INPUT
	WMODULETYPE : UINT;
	DWINSTANCE : UDINT;
	PCONNECTOR : POINTER TO IoConfigConnector;
END_VAR
END_METHOD

(* ---- L_ETCSLAVE_S131.pou ---- *)
FUNCTION_BLOCK L_ETCSLAVE_S131 EXTENDS L_ETCSlave
VAR
	HEVENTUPDATECONFIGURATIONDONE : RTS_IEC_HANDLE;
	HINTERFACEUPDATECONFIGURATIONDONE : RTS_IEC_HANDLE;
	ITFCALLBACK : CmpEventMgr.ICmpEventCallback;
	MYCONNECTOR : POINTER TO IoConfigConnector;
	SOWNCOMMPATH : STRING(199);
	WMODULECOUNT : WORD;
	IIOSLICES : ARRAY [1..c_MaxModules] OF POINTER TO L_IOSlice;
	FBS131_DIAGNOSTICS : L_ECC_S131_Diagnostics;
	C_MAXMODULES : WORD := 64;
END_VAR
END_FUNCTION_BLOCK

METHOD CHILDISIOSLICE : BOOL
VAR_INPUT
	PCHILD : POINTER TO IoConfigConnector;
END_VAR
END_METHOD

METHOD CYCLICCALL : UDINT
END_METHOD

METHOD EVENTCALLBACK : UDINT
VAR_INPUT
	PEVENTPARAM : POINTER TO EventParam;
END_VAR
END_METHOD

METHOD FB_EXIT : BOOL
VAR_INPUT
	BINCOPYCODE : BOOL;
END_VAR
END_METHOD

METHOD FB_INIT : BOOL
VAR_INPUT
	BINITRETAINS : BOOL;
	BINCOPYCODE : BOOL;
END_VAR
END_METHOD

METHOD GETIOSLICEINSTANCE : POINTER TO L_IOSlice
VAR_INPUT
	PCHILD_IOSLICE : POINTER TO IoConfigConnector;
END_VAR
END_METHOD

METHOD GETIOSLICES : BOOL
END_METHOD

METHOD INITIALIZE : UDINT
VAR_INPUT
	WMODULETYPE : UINT;
	DWINSTANCE : UDINT;
	PCONNECTOR : POINTER TO IoConfigConnector;
END_VAR
END_METHOD

METHOD READOWNCOMMPATH : BOOL
END_METHOD

METHOD REGISTERIOSLICE : BOOL
VAR_INPUT
	PSCIOSLICE : POINTER TO L_IOSlice;
	BYSLOTNUMBER : BYTE;
END_VAR
END_METHOD

METHOD WRITEDIAGINSTANCEADDRESS : BOOL
VAR_INPUT
	PCONNECTOR : POINTER TO IoConfigConnector;
END_VAR
END_METHOD

(* ---- L_ETCSLAVE_SAFETY.pou ---- *)
FUNCTION_BLOCK L_ETCSLAVE_SAFETY EXTENDS ETCSlave
VAR_OUTPUT
	PETCSLAVE : POINTER TO ETCSlave;
END_VAR
VAR
	ETCSLAVE : REFERENCE TO ETCSlave;
	FBSAFETYDIAGNOSTICS : L_ECC_Safety_Diagnostics;
END_VAR
END_FUNCTION_BLOCK

METHOD FB_EXIT : BOOL
VAR_INPUT
	BINCOPYCODE : BOOL;
END_VAR
END_METHOD

METHOD FB_INIT : BOOL
VAR_INPUT
	BINITRETAINS : BOOL;
	BINCOPYCODE : BOOL;
END_VAR
END_METHOD

METHOD INITIALIZE : UDINT
VAR_INPUT
	WMODULETYPE : UINT;
	DWINSTANCE : UDINT;
	PCONNECTOR : POINTER TO IoConfigConnector;
END_VAR
END_METHOD

METHOD WRITEDIAGINSTANCEADDRESS : BOOL
VAR_INPUT
	PCONNECTOR : POINTER TO IoConfigConnector;
END_VAR
END_METHOD

METHOD FB_REINIT : BOOL
END_METHOD

(* ---- L_IOSLICE.pou ---- *)
FUNCTION_BLOCK L_IOSLICE
VAR
	MODULEHANDLERBASE : L_IMHP_ModuleHandler := STRUCT(CompActiveDefault := TRUE, Layer := L_IMHP_Layer.Communication, CompType := L_IMHP_ComponentType.EtherCATSlave, DefaultRelationship := L_IMHP_RelationshipID.CommunicationView);
	MODULEID : L_ECC_eDeviceType;
	UIACTUALERROR : UINT;
	REGISTERONCOMPONENTDIRECTORY : L_IC1P_RegisterOnComponentDirectory;
	MYWMODULETYPE : UINT;
	MYDWINSTANCE : UDINT;
	MYPCONNECTOR : POINTER TO IoConfigConnector;
	MODULEHANDLER : L_IMHP_IModuleHandler;
END_VAR
END_FUNCTION_BLOCK

METHOD FB_INIT : BOOL
VAR_INPUT
	BINITRETAINS : BOOL;
	BINCOPYCODE : BOOL;
END_VAR
END_METHOD

METHOD INITIALIZE : UDINT
VAR_INPUT
	WMODULETYPE : UINT;
	DWINSTANCE : UDINT;
	PCONNECTOR : POINTER TO IoConfigConnector;
END_VAR
END_METHOD

METHOD READMODULEID : BOOL
VAR_INPUT
	PCONNECTOR : POINTER TO IoConfigConnector;
END_VAR
END_METHOD

METHOD WRITEINSTANCEADDRESS : BOOL
VAR_INPUT
	PCONNECTOR : POINTER TO IoConfigConnector;
END_VAR
END_METHOD

METHOD MDIAGNOSTICERRORTOERRORCODE : UINT
VAR_INPUT
	EDEVICETYPE : L_ECC_eDeviceType;
	DWERRORID : DWORD := 0;
END_VAR
END_METHOD

METHOD MERRORHANDLER : BOOL
VAR_INPUT
	ESEVERITY : _L_ECC_eSeverity := _L_ECC_eSeverity.Fault_Log;
	DWERRORID : DWORD := 0;
	WTEXTREFID : WORD;
END_VAR
END_METHOD

METHOD MSETCOMMPATH : BOOL
VAR_INPUT
	SPATH : STRING(199);
END_VAR
END_METHOD

(* ---- L_SUDP_PRMFILE_READWRITE_ETC.pou ---- *)
FUNCTION_BLOCK L_SUDP_PRMFILE_READWRITE_ETC EXTENDS L_SUDP_PRMFile_ReadWrite
VAR
	SDORD : L_ETC_CoE_SdoRead;
	FILESIZECHANGED : BOOL;
END_VAR
END_FUNCTION_BLOCK

METHOD BEFORESTARTEXECUTION
END_METHOD

METHOD READVALUEFROMFIELDBUS_LOOP : INT
END_METHOD

METHOD READVALUEFROMFIELDBUS_START
VAR_INPUT
	PARAMHDR : POINTER TO L_SUDP.L_SUDP_PARM_HDR;
	PBYBUFFER : POINTER TO BYTE;
	SZBUFFERSIZE : UINT;
END_VAR
END_METHOD
